{attribute 'qualified_only'}
{attribute 'strict'}
TYPE E_ConveyorState :
(
	IDLE,
    RUNNING,
	WAIT_EXIT,
    FAULT
);
END_TYPE

(* stored: Version 1.1.0.1, ProductVersion 3.1.4024.16
   DUT E_ConveyorState: Id {a4059b68-67bf-4031-9ea8-5deefe11b000} *)
